(*
1) This is the first item in the list.

   (a) This is the first subitem (1a).
   (b) This is the second subitem (1b).

2) This is the second item in the list.

   (a) This is the first subitem (2a).
   (b) This is the second subitem (2b).

#) This item is auto-enumerated.
*)

FUNCTION_BLOCK FB_Libdoc_OrderedNumberedEnumerationList
VAR_INPUT
    nVarA : INT;
    nVarB : INT;
END_VAR
VAR_OUTPUT
    nSum : INT;
END_VAR
VAR
END_VAR

END_FUNCTION_BLOCK

(* stored: Version 1.1.0.1, ProductVersion 3.1.4022.17
   POU FB_Libdoc_OrderedNumberedEnumerationList: Id {0b69690e-3bd4-4925-997e-bf4fd3f61cfd}, SpecialFunc None *)
